FUNCTION_BLOCK fbfalltrig
VAR_INPUT
	clkin:BOOL;
	
END_VAR
VAR_OUTPUT
	clkout:BOOL;
	
END_VAR
VAR
	bprevclk:BOOL;
	
END_VAR

clkout:= NOT clkin AND bprevclk;
bprevclk:=clkin;

END_FUNCTION_BLOCK

(* stored: Version 1.1.0.1, ProductVersion 3.1.4024.16
   POU fbfalltrig: Id {aa44cdb1-efb5-4aa3-9f13-bf47ea35e6a2}, SpecialFunc None *)
